SUBAPPLICATION ein (* Subapplication Type *)
  (* Standard: 61499-2 *)
  (* Version 1.0, 2023-02-07, franz *)
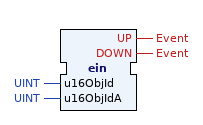
  EVENT_OUTPUT
    UP;
    DOWN;
  END_EVENT
  VAR_INPUT
    u16ObjId : UINT;
    u16ObjIdA : UINT;
  END_VAR
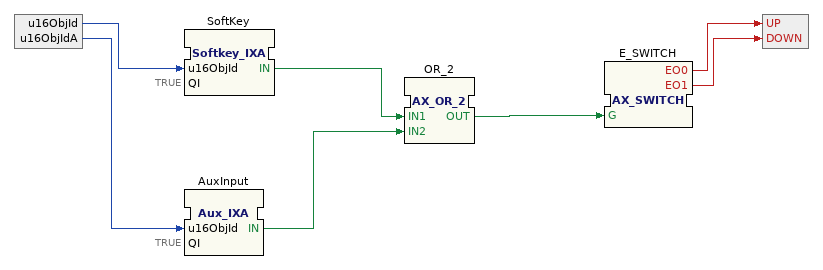
  FBS
    SoftKey : isobus::UT::io::Softkey::Softkey_IXA(QI := TRUE);
    AuxInput : isobus::UT::io::Auxiliary::IN::Aux_IXA(QI := TRUE);
    OR_2 : adapter::booleanOperators::AX_OR_2;
    E_SWITCH : adapter::events::unidirectional::AX_SWITCH;
  END_FBS
  EVENT_CONNECTIONS
    E_SWITCH.EO0 TO UP;
    E_SWITCH.EO1 TO DOWN;
  END_CONNECTIONS
  DATA_CONNECTIONS
    u16ObjIdA TO AuxInput.u16ObjId;
    u16ObjId TO SoftKey.u16ObjId;
  END_CONNECTIONS
  ADAPTER_CONNECTIONS
    SoftKey.IN TO OR_2.IN1;
    AuxInput.IN TO OR_2.IN2;
    OR_2.OUT TO E_SWITCH.G;
  END_CONNECTIONS
END_SUBAPPLICATION
